TYPE (* logiBUS_ENC Struct *)
  (* Version 1.0, 2026-11-26, Franz Höpfinger, initial API and implementation and/or initial documentation *)
  PACKAGE logiBUS::io::ENC;
  logiBUS_ENC_S : STRUCT
    Pin : USINT := 255;
  END_STRUCT;
END_TYPE
